(* IEC 61131-3 sources: llm-plc-st-eval/data/definitivo/gemini-3.1-pro-preview/A1/zero_shot, 3 files *)

(* ---- ejec_1.st ---- *)
```iecst
FUNCTION_BLOCK FB_PID
VAR_INPUT
    SP : REAL;      // Consigna (Setpoint)
    PV : REAL;      // Variable de proceso (Process Variable)
    Kp : REAL;      // Ganancia proporcional
    Ti : REAL;      // Tiempo integral (segundos)
    Td : REAL;      // Tiempo derivativo (segundos)
    ciclo : TIME;   // Período de muestreo
END_VAR

VAR_OUTPUT
    CV : REAL;      // Variable de control (0.0 a 100.0 %)
END_VAR

VAR
    e : REAL;                   // Error actual
    e_prev : REAL := 0.0;       // Error del ciclo anterior
    integral_sum : REAL := 0.0; // Sumatoria de la integral del error
    dt : REAL;                  // Tiempo de ciclo en segundos
    P_term : REAL;              // Término proporcional
    I_term : REAL;              // Término integral
    D_term : REAL;              // Término derivativo
    CV_pre : REAL;              // Salida preliminar para evaluar saturación
    CV_raw : REAL;              // Salida calculada sin limitar
END_VAR

// Convertir el tiempo de ciclo a segundos
dt := TIME_TO_REAL(ciclo) / 1000.0;

// Cálculo del error (salida aumenta si PV < SP)
e := SP - PV;

// Cálculo del término proporcional
P_term := Kp * e;

// Cálculo del término derivativo (sobre el error)
IF dt > 0.0 THEN
    D_term := Kp * Td * (e - e_prev) / dt;
ELSE
    D_term := 0.0;
END_IF;

// Cálculo del término integral y Anti-windup (Clamping)
IF Ti > 0.0 THEN
    // Calcular salida preliminar con la integral del ciclo anterior
    I_term := (Kp / Ti) * integral_sum;
    CV_pre := P_term + I_term + D_term;

    // Anti-windup: evitar acumular error si la salida está saturada en la misma dirección
    IF (CV_pre >= 100.0 AND e > 0.0) OR (CV_pre <= 0.0 AND e < 0.0) THEN
        // No se acumula el error (Clamping activo)
    ELSE
        // Se acumula el error en la integral
        IF dt > 0.0 THEN
            integral_sum := integral_sum + (e * dt);
        END_IF;
    END_IF;

    // Recalcular el término integral con el valor actualizado
    I_term := (Kp / Ti) * integral_sum;
ELSE
    // Desactivar acción integral si Ti <= 0.0
    integral_sum := 0.0;
    I_term := 0.0;
END_IF;

// Suma total de la ecuación PID estándar
CV_raw := P_term + I_term + D_term;

// Limitación de la salida (0.0 a 100.0)
IF CV_raw > 100.0 THEN
    CV := 100.0;
ELSIF CV_raw < 0.0 THEN
    CV := 0.0;
ELSE
    CV := CV_raw;
END_IF;

// Actualizar el error para el cálculo derivativo del próximo ciclo
e_prev := e;

END_FUNCTION_BLOCK
```

(* ---- ejec_2.st ---- *)
```iecst
FUNCTION_BLOCK FB_PID
VAR_INPUT
    SP : REAL;      // Consigna (Setpoint)
    PV : REAL;      // Variable de proceso
    Kp : REAL;      // Ganancia proporcional
    Ti : REAL;      // Tiempo integral (segundos)
    Td : REAL;      // Tiempo derivativo (segundos)
    ciclo : TIME;   // Período de muestreo
END_VAR

VAR_OUTPUT
    CV : REAL;      // Variable de control (0.0 a 100.0 %)
END_VAR

VAR
    e : REAL;           // Error actual
    e_prev : REAL;      // Error del ciclo anterior
    de_dt : REAL;       // Derivada del error
    dt : REAL;          // Tiempo de ciclo en segundos
    I_sum : REAL;       // Sumatoria de la integral del error
    I_new : REAL;       // Valor tentativo de la integral
    CV_tentative : REAL;// Salida tentativa para evaluar saturación
END_VAR

// Convertir tiempo de ciclo a segundos (REAL)
dt := TIME_TO_REAL(ciclo) / 1000.0;

// Evitar división por cero si el tiempo de ciclo es muy pequeño o cero
IF dt <= 0.0 THEN
    dt := 0.001;
END_IF;

// Cálculo del error (Acción directa: CV aumenta si PV < SP)
e := SP - PV;

// Cálculo de la derivada del error
de_dt := (e - e_prev) / dt;

// Acción Integral con Anti-windup (Clamping)
IF Ti > 0.0 THEN
    // Calcular integral tentativa
    I_new := I_sum + (e * dt);

    // Calcular salida tentativa para evaluar saturación
    CV_tentative := Kp * (e + (I_new / Ti) + (Td * de_dt));

    // Lógica de Clamping: evitar acumulación si satura en la misma dirección del error
    IF (CV_tentative >= 100.0 AND e > 0.0) OR (CV_tentative <= 0.0 AND e < 0.0) THEN
        // No se actualiza I_sum (se congela la integral)
    ELSE
        I_sum := I_new; // Se actualiza la integral
    END_IF;
ELSE
    I_sum := 0.0; // Desactivar acción integral si Ti <= 0.0
END_IF;

// Cálculo de la salida final (CV) antes de límites
IF Ti > 0.0 THEN
    CV := Kp * (e + (I_sum / Ti) + (Td * de_dt));
ELSE
    CV := Kp * (e + (Td * de_dt));
END_IF;

// Limitar la salida al rango 0.0 - 100.0 %
IF CV > 100.0 THEN
    CV := 100.0;
ELSIF CV < 0.0 THEN
    CV := 0.0;
END_IF;

// Guardar el error actual para el cálculo derivativo del próximo ciclo
e_prev := e;

END_FUNCTION_BLOCK
```

(* ---- ejec_3.st ---- *)
```iecst
FUNCTION_BLOCK FB_PID
VAR_INPUT
    SP : REAL;      (* Consigna (Setpoint) *)
    PV : REAL;      (* Variable de proceso *)
    Kp : REAL;      (* Ganancia proporcional *)
    Ti : REAL;      (* Tiempo integral en segundos *)
    Td : REAL;      (* Tiempo derivativo en segundos *)
    ciclo : TIME;   (* Período de muestreo *)
END_VAR

VAR_OUTPUT
    CV : REAL;      (* Variable de control (0.0 a 100.0) *)
END_VAR

VAR
    e : REAL;       (* Error actual *)
    e_prev : REAL;  (* Error del ciclo anterior *)
    I_term : REAL;  (* Término integral acumulado *)
    P_term : REAL;  (* Término proporcional *)
    D_term : REAL;  (* Término derivativo *)
    dt : REAL;      (* Tiempo de ciclo en segundos *)
END_VAR

(* Convertir el tiempo de ciclo a segundos (REAL) *)
dt := TIME_TO_REAL(ciclo) / 1000.0;

(* Evitar ejecución si el tiempo de ciclo es inválido o cero *)
IF dt > 0.0 THEN

    (* Cálculo del error (Acción directa: si PV < SP, e > 0 y CV aumenta) *)
    e := SP - PV;

    (* 1. Término Proporcional *)
    P_term := Kp * e;

    (* 2. Término Integral con Anti-windup (Clamping) *)
    IF Ti > 0.0 THEN
        (* Evaluar saturación de la salida en el ciclo anterior y el signo del error *)
        IF NOT ((CV >= 100.0 AND e > 0.0) OR (CV <= 0.0 AND e < 0.0)) THEN
            I_term := I_term + (Kp * e * dt) / Ti;
        END_IF;
    ELSE
        (* Desactivar acción integral si Ti <= 0.0 *)
        I_term := 0.0;
    END_IF;

    (* 3. Término Derivativo (calculado sobre el error) *)
    D_term := Kp * Td * (e - e_prev) / dt;

    (* Actualizar el error para el cálculo derivativo del próximo ciclo *)
    e_prev := e;

    (* Cálculo de la salida total *)
    CV := P_term + I_term + D_term;

    (* Limitación de la salida (Saturación 0.0 a 100.0) *)
    IF CV > 100.0 THEN
        CV := 100.0;
    ELSIF CV < 0.0 THEN
        CV := 0.0;
    END_IF;

END_IF;
END_FUNCTION_BLOCK
```
